(* IEC 61131-3 sources: plc-process-lib/src/Interfaces/I_Device, 1 file *)

(* ---- RequestMode.method.decl.st ---- *)
// Запрос режима: Auto, Manual, OutOfService — как команда stCmd; Local и прочее — FALSE.
// Имя параметра не eMode: оно затенило бы переменную базы (L3)
METHOD RequestMode : BOOL
VAR_INPUT
    eNewMode : E_DeviceMode;   // требуемый режим
END_VAR
